FUNCTION_BLOCK AD2_D_TO_DWORD (* Composite FB for convert AD2 to DWORD *)
  (* Standard: 61499-2; Description: Copyright (c) 2026 HR Agrartechnik GmbH This program and the accompanying materials are made available under the terms of the Eclipse Public License 2.0 which is available at https://www.eclipse.org/legal/epl-2.0/ SPDX-License-Identifier: EPL-2.0 *)
  (* Version 1.0, 2026-11-13, Franz Höpfinger, HR Agrartechnik GmbH, Initial Version - Luecke geschlossen (analog zu AB2_B_TO_BYTE) *)
  PACKAGE adapter::conversion::bidirectional;
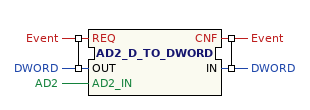
  EVENT_INPUT
    REQ WITH OUT; (* Request to Adapter *)
  END_EVENT
  EVENT_OUTPUT
    CNF WITH IN; (* Confirmation from Adapter *)
  END_EVENT
  VAR_INPUT
    OUT : DWORD; (* Output data to Adapter *)
  END_VAR
  VAR_OUTPUT
    IN : DWORD; (* Input data from Adapter *)
  END_VAR
  SOCKETS
    AD2_IN : adapter::types::bidirectional::AD2; (* Adapter Input *)
  END_SOCKETS
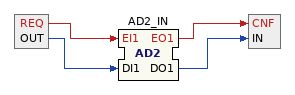
  EVENT_CONNECTIONS
    AD2_IN.EO1 TO CNF;
    REQ TO AD2_IN.EI1;
  END_CONNECTIONS
  DATA_CONNECTIONS
    AD2_IN.DO1 TO IN;
    OUT TO AD2_IN.DI1;
  END_CONNECTIONS
END_FUNCTION_BLOCK
